KUKA KRL data list: bt_cell.dat

&ACCESS RVP
&REL 1
&COMMENT bt2krl sim job loop data plan 16#4F80
DEFDAT BT_CELL
   ; Generated by bt2krl 0.1.0 from bt2plc plan bt_1792076124_welding_cell_2_small (cell welding_cell_2_small), PLAN_ID 16#4F80
   ; Robot robot2 (R2), controller robot2, model KR240R2900_ULTRA, joint mapping identity
   ; Profile sim (bt2plc simulator telegram). NEVER install on a VW KS24 robot:
   ; its signals collide with the VW standard (Fertigmeldung, interlocks, PRG_NR).
   ; Do not edit: regenerate with bt2krl (plain KRL, no inline forms).
ENDDAT
